Fanuc KAREL source: kc00002.KL

-- PROVISIONAL review KL for V770-1; original PC SHA256 c7362087b31b84d8b9767280304104a050437004b46a1f6e58b1fecc39624dbe
-- Incomplete behavior may be omitted. Consult companion uncertainty JSON. Do not deploy.
PROGRAM KC00002
%NOLOCKGROUP
BEGIN
  -- UNRESOLVED_PC offsets 5-33; opcodes 27,22,22,22,22,31
  -- UNRESOLVED_PC offsets 38-42; opcodes 7F
END KC00002
